TYPE "FRK_ConfigInteger"
VERSION : 0.1
   STRUCT
      "Used" {ExternalAccessible := 'False'; ExternalVisible := 'False'; ExternalWritable := 'False'} : Int;
      "Limbs" {ExternalAccessible := 'False'; ExternalVisible := 'False'; ExternalWritable := 'False'} : Array[0..101] of UDInt;
   END_STRUCT;
END_TYPE
